TYPE ST_PolarIIChamber_AngularPositionParam :
STRUCT
	Position : LREAL; // deg
END_STRUCT
END_TYPE

(* stored: Version 1.1.0.1, ProductVersion 3.1.4026.18
   DUT ST_PolarIIChamber_AngularPositionParam: Id {14000000-0000-0000-0000-000000000078} *)
